// TIA Portal V21 export
// export: Created 2026-11-11T00:47:32.5415158Z, ExportSetting WithDefaults, DisplayName Totally Integrated Automation Portal, DisplayVersion V21 Update 3, DisplayName STEP 7 Professional, DisplayVersion V21 Update 3, DisplayName STEP 7 Safety, DisplayVersion V21, DisplayName Tech WebApplication, DisplayVersion V21, DisplayName WinCC Basic/Comfort/Advanced, DisplayVersion V21 Update 3, DisplayName WinCC Unified, DisplayVersion V21 Update 3
FUNCTION_BLOCK "FB_Fbd_ex124"   // FB134, FBD
{ S7_Optimized_Access := 'TRUE' }
VERSION : 0.1
// stored: AutoNumber true, IsIECCheckEnabled false, IsRetainMemResEnabled false, MemoryReserve 100, SetENOAutomatically false, UDAEnableTagReadback false
   VAR_OUTPUT
      v_ret_val : Int;
   END_VAR
   VAR_IN_OUT
      v_top_si : Array[0..99] of Byte;
      v_start_up_si : Array[0..99] of Byte;
   END_VAR
BEGIN

REGION Network 1: RD_SINFO - Read current OB start information
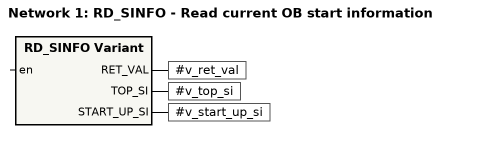
   #v_ret_val := RD_SINFO(TOP_SI => #v_top_si, START_UP_SI => #v_start_up_si);
END_REGION
END_FUNCTION_BLOCK
